// Core S3.12 - the MEASURE result, valid on Done.
TYPE ST_AnalogInputOutCmd :
STRUCT
    Value : LREAL;    // the measured value
END_STRUCT
END_TYPE

(* stored: Version 1.1.0.1, ProductVersion 3.1.4024.12
   DUT ST_AnalogInputOutCmd: Id {fcb69756-ad4a-490a-9b7f-532059b57287} *)
